(* IEC 61131-3 sources: openplc-editor-canopen/src/backend/shared/transpilers/st-transpiler/__tests__/fixtures/ld-relayout-corpus/ld-corpus-basic/expected-st, 4 files *)

(* ---- _project.st ---- *)
CONFIGURATION Config0

  RESOURCE Res0 ON PLC
    TASK task0(INTERVAL := T#20ms,PRIORITY := 1);
    PROGRAM instance0 WITH task0 : main;
  END_RESOURCE
END_CONFIGURATION

(* ---- Auxiliary.st ---- *)
PROGRAM Auxiliary
  VAR
    aux_a : BOOL;
    TON0 : TON;
    aux_x1 : BOOL;
    aux_x2 : BOOL;
    aux_x3 : BOOL;
    aux_et1 : TIME;
    aux_b : BOOL;
    CTU0 : CTU;
    aux_y1 : BOOL;
    aux_r2 : BOOL;
    aux_cv2 : INT;
    aux_c : BOOL;
    TOF0 : TOF;
    aux_z1 : BOOL;
    aux_z2 : BOOL;
    aux_d : BOOL;
    aux_e : BOOL;
    aux_w1 : BOOL;
  END_VAR

  TON0(IN := aux_a, PT := T#1s);
  aux_et1 := TON0.ET;
  aux_x1 := TON0.Q;
  aux_x2 := TON0.Q;
  aux_x3 := TON0.Q;
  CTU0(CU := aux_b, R := aux_r2, PV := 3);
  aux_y1 := CTU0.Q;
  aux_cv2 := CTU0.CV;
  TOF0(IN := aux_c OR aux_d, PT := T#2s);
  aux_z1 := TOF0.Q;
  aux_z2 := TOF0.Q;
  aux_w1 := aux_e;
END_PROGRAM

(* ---- Blocks.st ---- *)
PROGRAM Blocks
  VAR
    b03_enable : BOOL;
    TON0 : TON;
    b03_done : BOOL;
    b03_start : BOOL;
    b03_q : BOOL;
    b03_et : TIME;
    b04_up : BOOL;
    CTUD0 : CTUD;
    b04_at_max : BOOL;
    b04_down : BOOL;
    b04_reset : BOOL;
    b04_load : BOOL;
    b04_at_min : BOOL;
    b04_count : INT;
    b05_run : BOOL;
    ONTIME0 : ONTIME;
    b05_eno : BOOL;
    b05_in : BOOL;
    b05_rst : BOOL;
    b05_seconds : UDINT;
    b05_cycles : UDINT;
    b08_go : BOOL;
    TON1 : TON;
    b08_q : BOOL;
    b08_et : TIME;
    b09_go : BOOL;
    TON2 : TON;
    b09_eno : BOOL;
    b09_in : BOOL;
    b09_q : BOOL;
    b09_et : TIME;
  END_VAR

  TON0(EN := b03_enable, IN := b03_start, PT := T#2s);
  b03_done := TON0.ENO;
  IF TON0.ENO THEN
      b03_q := TON0.Q;
  END_IF;
  IF TON0.ENO THEN
      b03_et := TON0.ET;
  END_IF;
  CTUD0(CU := b04_up, CD := b04_down, R := b04_reset, LD := b04_load, PV := 20);
  b04_at_max := CTUD0.QU;
  b04_at_min := CTUD0.QD;
  b04_count := CTUD0.CV;
  ONTIME0(EN := b05_run, IN := b05_in, RST := b05_rst, SECONDS := b05_seconds, CYCLES := b05_cycles);
  b05_eno := ONTIME0.ENO;
  TON1(IN := b08_go, PT := T#500ms);
  b08_q := TON1.Q;
  b08_et := TON1.ET;
  TON2(EN := b09_go, IN := b09_in, PT := T#1s);
  b09_eno := TON2.ENO;
  IF TON2.ENO THEN
      b09_q := TON2.Q;
  END_IF;
  IF TON2.ENO THEN
      b09_et := TON2.ET;
  END_IF;
END_PROGRAM

(* ---- Main.st ---- *)
PROGRAM Main
  VAR
    b01_start : BOOL;
    b01_motor : BOOL;
    b01_permit : BOOL;
    b01_guard : BOOL;
    b02_a : BOOL;
    b02_out : BOOL;
    b02_b : BOOL;
    b02_c : BOOL;
    b02_e : BOOL;
    b06_run : BOOL;
    b06_lamp1 : BOOL;
    b06_lamp2 : BOOL;
    b06_lamp3 : BOOL;
    b07_cmd : BOOL;
    b07_latch : BOOL;
    b07_unlatch : BOOL;
    b07_rise : BOOL;
    b07_fall : BOOL;
    b11_conveyor_section_one_upstream_permissive_signal : BOOL;
    TON0 : TON;
    b11_conveyor_section_one_downstream_motor_run_command : BOOL;
    b11_conveyor_section_one_start_delay_preset_time_value : TIME;
    b11_conveyor_section_one_start_delay_elapsed_time_value : TIME;
    _TMP_R_TRIG1898394 : R_TRIG;
    _TMP_F_TRIG2000051 : F_TRIG;
  END_VAR

  b01_motor := b01_guard AND b01_permit AND b01_start;
  b02_out := b02_a OR b02_b OR b02_e AND b02_c;
  b06_lamp1 := b06_run;
  b06_lamp2 := b06_run;
  b06_lamp3 := b06_run;
  IF b07_cmd THEN
    b07_latch := TRUE; (*set*)
  END_IF;
  IF b07_cmd THEN
    b07_unlatch := FALSE; (*reset*)
  END_IF;
  _TMP_R_TRIG1898394(CLK := b07_cmd);
  b07_rise := _TMP_R_TRIG1898394.Q;
  _TMP_F_TRIG2000051(CLK := b07_cmd);
  b07_fall := _TMP_F_TRIG2000051.Q;
  TON0(IN := b11_conveyor_section_one_upstream_permissive_signal, PT := b11_conveyor_section_one_start_delay_preset_time_value);
  b11_conveyor_section_one_downstream_motor_run_command := TON0.Q;
  b11_conveyor_section_one_start_delay_elapsed_time_value := TON0.ET;
END_PROGRAM
